Fanuc KAREL source: kb00157.KL

-- PROVISIONAL review KL for V940-1; original PC SHA256 6c1dd87d78f99e8e683ced23950ad856c55b9fb189b482805e2f5418ac2971b6
-- Incomplete behavior may be omitted. Consult companion uncertainty JSON. Do not deploy.
PROGRAM KB00157
%NOLOCKGROUP
BEGIN
  -- V9_ZERO_TABLE_METADATA_HINT layout=0002_ascii; no indexed target words; source/name/runtime held
  -- UNRESOLVED_PC offsets 5-12; opcodes 9D,23
  -- UNRESOLVED_PC offsets 17-33; opcodes 27,22,31,23
  -- UNRESOLVED_PC offsets 38-42; opcodes 7F
END KB00157
